FUNCTION_BLOCK TcoKukaKss_StopMovementsAndProgramTask_v_9_3_x EXTENDS TcoKukaKssTask_v_9_3_x
VAR
	_stopType : TcoAbstractions.eTcoRoboticsStopType;
END_VAR

IF Execute() THEN
	_blink(inOnTime:=T#500MS,inOffTime:=T#500MS);

	IF _progress = 0 THEN
		IF CheckReferences() THEN
			_progress := _progress + 1;
		END_IF
	END_IF

	IF _progress = 1 THEN
		// AX step 0: waiting for 'RobotStopped'
		inoControl.MoveEnable := FALSE;
		_varInfo :=__VARINFO(inoStatus.State.RobotStopped);
		THIS^.Messenger.OnCondition(_infoTimer.Q AND NOT inoStatus.State.RobotStopped).Warning(_sb.Clear().Append('<#Waiting for signal: #>').Append(_varInfo.Symbol).ToString());
		IF inoStatus.State.RobotStopped THEN
			_progress := _progress + 1;
		END_IF
	END_IF

	IF _progress = 2 THEN
		// AX step 1: waiting for 'ProActive' to be off
		_varInfo :=__VARINFO(inoStatus.State.ProActive);
		THIS^.Messenger.OnCondition(_infoTimer.Q AND inoStatus.State.ProActive).Warning(_sb.Clear().Append('<#Waiting for signal: #>').Append(_varInfo.Symbol).Append('<# is OFF#>').ToString());
		IF NOT inoStatus.State.ProActive THEN
			_progress := _progress + 1;
		END_IF
	END_IF

	IF _progress = 3 THEN
		DoneWhen(TRUE);
	END_IF

	CallTimers(TRUE);
	THIS^.ThrowWhen(_errorTimer.Q);
END_IF

IF THIS^.Error AND NOT _errorMessage.Pinned THEN
	THIS^.Restore();
END_IF

METHOD INTERNAL InvokeWithParams : ITcoTaskStatus
VAR_INPUT
	inStopType : eTcoRoboticsStopType;
END_VAR
_stopType := inStopType;
InvokeWithParams := THIS^.Invoke();
END_METHOD

METHOD PUBLIC FB_init : BOOL
VAR_INPUT
    bInitRetains : BOOL; // if TRUE, the retain variables are initialized (warm start / cold start)
    bInCopyCode : BOOL; // if TRUE, the instance afterwards gets moved into the copy code (online change)
    ParentObject : ITcoObject;
END_VAR
END_METHOD

(*~
	<docu>
		<summary>
			Executes when task is aborted.
		</summary>			
	</docu>	
~*)
METHOD PROTECTED OnAbort
IF __ISVALIDREF(inoStatus) THEN THIS^.inoStatus.ActionDescription := '<#Stop movements and program was aborted.#>'; END_IF;
END_METHOD

(*~
	<docu>
		<summary>
			Executes when task reaches the ```Done``` state .
		</summary>			
	</docu>	
~*)
METHOD PROTECTED OnDone
IF __ISVALIDREF(inoStatus) THEN THIS^.inoStatus.ActionDescription := '<#Stop movements and program finished successfully.#>'; END_IF;
_progress := 0;
END_METHOD

(*~
	<docu>
		<summary>
			Executes when task reaches the ```Error``` state.
		</summary>			
	</docu>	
~*)
METHOD PROTECTED OnError
VAR
	description: STRING;
END_VAR
description := '<#Stop movements and program finished with error.#>';
IF __ISVALIDREF(inoStatus) THEN THIS^.inoStatus.ActionDescription := description; END_IF;
THIS^._errorMessage.Error(_sb.Clear().Append(description).Append(' To restore acknowledge this alarm.').ToString()).Pin();
END_METHOD

METHOD PROTECTED OnStart
IF __ISVALIDREF(inoStatus) THEN THIS^.inoStatus.ActionDescription := '<#Stop movements and program started.#>'; END_IF;
CallTimers(FALSE);
END_METHOD

(*~
	<docu>
		<summary>
			Restores this instance to the Ready state. Can be called explicitly or from within one of the restore mechanisms.
			<para>
				See also <see cref="PlcDocu.TcoCore.TcoTask.AutoRestorable()"/>
			</para>
		</summary>
	</docu>
~*)
METHOD Restore : ITcoRestorable
SUPER^.Restore();
END_METHOD

END_FUNCTION_BLOCK

(* stored: Version 1.1.0.1, ProductVersion 3.1.4024.12
   POU TcoKukaKss_StopMovementsAndProgramTask_v_9_3_x: Id {4ecaa873-4379-4a61-a3dc-249a6038f264}, SpecialFunc None
   Method InvokeWithParams: Id {90e1d21f-2fdd-45e2-b8bb-47356c40529d}
   Method FB_init: Id {c991eb92-1b08-434a-82fb-12adb347620b}
   Method OnAbort: Id {3701f0f8-63c8-402b-a9de-48c046d10342}
   Method OnDone: Id {cce8d677-1db0-4dbe-8398-dab7cf10148a}
   Method OnError: Id {c9a73734-15f2-4dcf-9b04-b928dc552e9a}
   Method OnStart: Id {2ea2d78f-f7aa-4292-953a-95c64b2974ef}
   Method Restore: Id {94375718-3eb2-47c8-86be-ed372d2efc1a} *)
